// TIA Portal V21 export
Screen "T01_Rect"  1024x768, Number=21
  ScreenLayer 
    Rectangle "P_CellRect" at 0,0 size 100x30
